FUNCTION_BLOCK T_E_text_MainControl EXTENDS KOSTAL_AF2024_Core_Text.T_E_Text
VAR
END_VAR

PROPERTY busy : KOSTAL_AF2024_Core_Text.ST_E_Text
GET
busy.Number:= 36;
END_GET
END_PROPERTY

PROPERTY lastCycle : KOSTAL_AF2024_Core_Text.ST_E_Text
GET
lastCycle.Number:= 37;
END_GET
END_PROPERTY

PROPERTY name : KOSTAL_AF2024_Core_Text.ST_E_Text
GET
name.Number:= 2;
END_GET
END_PROPERTY

PROPERTY nextPage : KOSTAL_AF2024_Core_Text.ST_E_Text
GET
nextPage.Number:= 61;
END_GET
END_PROPERTY

PROPERTY off : KOSTAL_AF2024_Core_Text.ST_E_Text
GET
off.Source:= KOSTAL_AF2024_Core_Text.E_Source.Common;
off.Number:= 2;
END_GET
END_PROPERTY

PROPERTY onToHomeReleased : KOSTAL_AF2024_Core_Text.ST_E_Text
GET
onToHomeReleased.Source:= KOSTAL_AF2024_Core_Text.E_Source.Common;
onToHomeReleased.Number:= 42;
END_GET
END_PROPERTY

PROPERTY onWith_0 : KOSTAL_AF2024_Core_Text.ST_E_Text
GET
onWith_0.Source:= KOSTAL_AF2024_Core_Text.E_Source.Common;
onWith_0.Number:= 65;
END_GET
END_PROPERTY

PROPERTY participantNotReady : KOSTAL_AF2024_Core_Text.ST_E_Text
GET
participantNotReady.Number:= 12;
END_GET
END_PROPERTY

PROPERTY powerOn : KOSTAL_AF2024_Core_Text.ST_E_Text
GET
powerOn.Number:= 44;
END_GET
END_PROPERTY

PROPERTY previousPage : KOSTAL_AF2024_Core_Text.ST_E_Text
GET
previousPage.Number:= 60;
END_GET
END_PROPERTY

PROPERTY readyToStart : KOSTAL_AF2024_Core_Text.ST_E_Text
GET
readyToStart.Number:=35;
END_GET
END_PROPERTY

PROPERTY refresh : KOSTAL_AF2024_Core_Text.ST_E_Text
GET
refresh.Number:= 62;
END_GET
END_PROPERTY

PROPERTY reset : KOSTAL_AF2024_Core_Text.ST_E_Text
GET
reset.Source:= Kostal_AF2024_Core_Text.E_Source.Common;
reset.Number:= 7;
END_GET
END_PROPERTY

PROPERTY run : KOSTAL_AF2024_Core_Text.ST_E_Text
GET
run.Number:= 5;
END_GET
END_PROPERTY

PROPERTY safetyInError : KOSTAL_AF2024_Core_Text.ST_E_Text
GET
safetyInError.Number:= 30;
END_GET
END_PROPERTY

PROPERTY setAutomaticMode : KOSTAL_AF2024_Core_Text.ST_E_Text
GET
setAutomaticMode.Number:=41;
END_GET
END_PROPERTY

PROPERTY setManualMode : KOSTAL_AF2024_Core_Text.ST_E_Text
GET
setManualMode.Number:= 40;
END_GET
END_PROPERTY

PROPERTY start : KOSTAL_AF2024_Core_Text.ST_E_Text
GET
start.Source:= KOSTAL_AF2024_Core_Text.E_Source.Common;
start.Number:= 5;
END_GET
END_PROPERTY

PROPERTY step_0_actual_1 : KOSTAL_AF2024_Core_Text.ST_E_Text
GET
step_0_actual_1.Source:= KOSTAL_AF2024_Core_Text.E_Source.Common;
step_0_actual_1.Number:= 11;
END_GET
END_PROPERTY

PROPERTY step_0_doesNotExist : KOSTAL_AF2024_Core_Text.ST_E_Text
GET
step_0_doesNotExist.Source:= KOSTAL_AF2024_Core_Text.E_Source.Common;
step_0_doesNotExist.Number:= 12;
END_GET
END_PROPERTY

PROPERTY stop : KOSTAL_AF2024_Core_Text.ST_E_Text
GET
stop.Source:= KOSTAL_AF2024_Core_Text.E_Source.Common;
stop.Number:= 4;
END_GET
END_PROPERTY

PROPERTY textHandlerIsNotReady : KOSTAL_AF2024_Core_Text.ST_E_Text
GET
textHandlerIsNotReady.Source:= KOSTAL_AF2024_Core_Text.E_Source.Common;
textHandlerIsNotReady.Number:= 20;
END_GET
END_PROPERTY

PROPERTY waitForAirPressure_0_1_2 : KOSTAL_AF2024_Core_Text.ST_E_Text
GET
waitForAirPressure_0_1_2.Number:= 31;
END_GET
END_PROPERTY

PROPERTY waitForAllOff : KOSTAL_AF2024_Core_Text.ST_E_Text
GET
waitForAllOff.Number:= 10;
END_GET
END_PROPERTY

PROPERTY waitForAllOn : KOSTAL_AF2024_Core_Text.ST_E_Text
GET
waitForAllOn.Number:= 11;
END_GET
END_PROPERTY

PROPERTY waitForPowerOn : KOSTAL_AF2024_Core_Text.ST_E_Text
GET
waitForPowerOn.Number:= 13;
END_GET
END_PROPERTY

PROPERTY waitFromHome : KOSTAL_AF2024_Core_Text.ST_E_Text
GET
waitFromHome.Number:= 43;
END_GET
END_PROPERTY

END_FUNCTION_BLOCK

(* stored: Version 1.1.0.1, ProductVersion 3.1.4024.12
   POU T_E_text_MainControl: Id {846e043b-cd09-4e3b-97f9-17b4385cca23}, SpecialFunc None
   Property busy: Id {f2e16b16-5d64-48c2-af31-ab14913a4587}
   Get Get: Id {d4012105-90ac-4e02-8417-8f1afc872b64}
   Property lastCycle: Id {295bd6f6-f4a7-4426-8c1c-5793400fbf32}
   Get Get: Id {d025d58a-8bcd-498b-ad76-708ac6324dab}
   Property name: Id {da5fa430-5ab5-40ef-ad4e-f848c2e3231c}
   Get Get: Id {21698cef-9f1a-4c1b-80bf-c8a317a0df5d}
   Property nextPage: Id {160deb59-0252-40cf-82cf-b6c5f428fa65}
   Get Get: Id {6223458b-7941-4e6a-a113-f0e00a2bc9f3}
   Property off: Id {5d9478bb-aa0f-4983-be74-9bf0ff6a259f}
   Get Get: Id {c99538f7-0a3b-4a6e-9b86-aab097fc9648}
   Property onToHomeReleased: Id {d4fd038c-122a-4416-a234-85b79803d1bf}
   Get Get: Id {9bf12418-bb17-4610-9115-0449fd3668d2}
   Property onWith_0: Id {aa112115-705d-4dce-8894-610fae71219f}
   Get Get: Id {1dc0401f-16ec-4458-a670-24be89555b14}
   Property participantNotReady: Id {164430b4-6585-4567-b676-f8f5bd8ab700}
   Get Get: Id {370f4149-82d8-4391-9e72-6fe9fff3683c}
   Property powerOn: Id {29cd478f-1b0a-4bc1-946f-5e81d45d43c5}
   Get Get: Id {9c3181a9-b276-4b40-8328-6659eb4d9189}
   Property previousPage: Id {70a6b168-cceb-4116-9e15-8317aaa1335d}
   Get Get: Id {44da14be-984e-424c-a552-2d61505dc0c9}
   Property readyToStart: Id {70c7c524-006f-4bf1-8877-089547d5a251}
   Get Get: Id {e1e7dfc6-6ba4-4ab1-8f6c-d70910afb434}
   Property refresh: Id {520478a6-8462-41df-ae2e-c4968714d56b}
   Get Get: Id {cefbc5d0-a054-4492-810c-b3b538afcc1d}
   Property reset: Id {ec0fa5f1-befe-4a6c-bf31-7ce4b7496dd2}
   Get Get: Id {8e879788-ea21-487d-b178-eac60b7078d6}
   Property run: Id {6be80cb1-547c-4c61-943b-d324be3d1206}
   Get Get: Id {e819674b-4d98-452d-948d-c5af1e53e9e7}
   Property safetyInError: Id {b230dc2b-c2f9-4a5b-9d3c-35c8e035ef53}
   Get Get: Id {852824af-83e3-4508-92b1-4afa75b3ba63}
   Property setAutomaticMode: Id {58b7c639-15b3-49d0-8b7d-ef309920785a}
   Get Get: Id {8972107c-e1de-46d1-b381-73d98ebdd627}
   Property setManualMode: Id {25a8c015-8502-4fce-90c5-611ad50f9eff}
   Get Get: Id {eabf2140-395b-49c0-bdf0-d58d3a15e389}
   Property start: Id {4b610585-bb79-4642-ab13-2091eea25464}
   Get Get: Id {d496ac44-22c9-4902-8d61-bc94dd29cef2}
   Property step_0_actual_1: Id {75a27154-3432-4ae3-beac-c01548651dd9}
   Get Get: Id {692bbf4d-dda4-40f8-8819-962b22a4dd4c}
   Property step_0_doesNotExist: Id {ea175b03-d17a-4bee-980b-39935bf162ba}
   Get Get: Id {397b4884-c0f6-4186-937d-8df6a114c254}
   Property stop: Id {27b4cf7d-6988-40f3-9263-e75321a3aa9d}
   Get Get: Id {180ae232-403d-4fa0-b985-e5aacf288930}
   Property textHandlerIsNotReady: Id {ae5da327-636d-483f-bcb1-60cccc96df8c}
   Get Get: Id {48a258c8-763a-47cb-82a7-bc899f987156}
   Property waitForAirPressure_0_1_2: Id {3daa9b1d-555b-4229-b0ac-4955befb6234}
   Get Get: Id {dd775d49-14eb-4904-8d56-fd60d467c36d}
   Property waitForAllOff: Id {3e548221-719d-4f6f-829f-46084fe6e905}
   Get Get: Id {fc257d21-3650-401e-914f-4cc259848e35}
   Property waitForAllOn: Id {0065be06-5385-46e2-8066-4311ebd14f92}
   Get Get: Id {009d783e-d9fd-451d-86c3-654d1c2bc66c}
   Property waitForPowerOn: Id {cec5138f-a579-4d3a-b92a-b6fcba67d54b}
   Get Get: Id {b8f843ec-76f6-4745-b767-d6b92ad5cb98}
   Property waitFromHome: Id {716dbd28-0c3a-4a3f-b61c-2a04cfb00672}
   Get Get: Id {e90f0f83-1e86-467c-bd59-6d6f4d6f1ed1} *)
